(* IEC 61131-3 sources: IEC61131-3_ST_SCL_Mutation_Generator/Tests/mutatedCode_multiple_breakers_management_H, 6 files *)

(* ---- M1399.st ---- *)
FUNCTION_BLOCK "FB_MotorControl"

VAR_INPUT
    Pressure_LOW : DINT;
END_VAR

VAR_OUTPUT
    Motor_Critical : BOOL;
END_VAR

VAR
    Threshold : DINT := 36464;
END_VAR

BEGIN

    IF Pressure_LOW > Threshold THEN (* MUTATED: REL_OP_REPLACE *)
        Motor_Critical := TRUE;
    ELSE
        Motor_Critical := FALSE;
    END_IF;

END_FUNCTION_BLOCK

(* ---- M1400.st ---- *)
FUNCTION_BLOCK "FB_MotorControl"

VAR_INPUT
    Pressure_LOW : DINT;
END_VAR

VAR_OUTPUT
    Motor_Critical : BOOL;
END_VAR

VAR
    Threshold : DINT := 36464;
END_VAR

BEGIN

    IF Pressure_LOW < Threshold THEN
        Motor_Critical := FALSE; (* MUTATED: BOOL_CONST_REPLACE *)
    ELSE
        Motor_Critical := FALSE;
    END_IF;

END_FUNCTION_BLOCK

(* ---- M1401.st ---- *)
FUNCTION_BLOCK "FB_MotorControl"

VAR_INPUT
    Pressure_LOW : DINT;
END_VAR

VAR_OUTPUT
    Motor_Critical : BOOL;
END_VAR

VAR
    Threshold : DINT := 36464;
END_VAR

BEGIN

    IF Pressure_LOW < Threshold THEN
        Motor_Critical := TRUE;
    ELSE
        Motor_Critical := TRUE; (* MUTATED: BOOL_CONST_REPLACE *)
    END_IF;

END_FUNCTION_BLOCK

(* ---- M1402.st ---- *)
FUNCTION_BLOCK "FB_MotorControl"

VAR_INPUT
    Pressure_LOW : DINT;
END_VAR

VAR_OUTPUT
    Motor_Critical : BOOL;
END_VAR

VAR
    Threshold : DINT := 36464;
END_VAR

BEGIN

    IF Pressure_LOW < Threshold THEN
        Motor_Critical := NOT (TRUE); (* MUTATED: ASSIGN_NEGATE *)
    ELSE
        Motor_Critical := FALSE;
    END_IF;

END_FUNCTION_BLOCK

(* ---- M1403.st ---- *)
FUNCTION_BLOCK "FB_MotorControl"

VAR_INPUT
    Pressure_LOW : DINT;
END_VAR

VAR_OUTPUT
    Motor_Critical : BOOL;
END_VAR

VAR
    Threshold : DINT := 36464;
END_VAR

BEGIN

    IF Pressure_LOW < Threshold THEN
        Motor_Critical := TRUE;
    ELSE
        Motor_Critical := NOT (FALSE); (* MUTATED: ASSIGN_NEGATE *)
    END_IF;

END_FUNCTION_BLOCK

(* ---- M1404.st ---- *)
FUNCTION_BLOCK "FB_MotorControl"

VAR_INPUT
    Pressure_LOW : DINT;
END_VAR

VAR_OUTPUT
    Motor_Critical : BOOL;
END_VAR

VAR
    Threshold : DINT := 36464;
END_VAR

BEGIN

    IF NOT (Pressure_LOW < Threshold) THEN (* MUTATED: COND_NEGATE *)
        Motor_Critical := TRUE;
    ELSE
        Motor_Critical := FALSE;
    END_IF;

END_FUNCTION_BLOCK
